Fanuc KAREL source: kt00489.KL

-- PROVISIONAL review KL for V1013-1; original PC SHA256 af2217d419cc08992401e6106b01a0b923f42a5de7de44bf260eaf8e4cc73e97
-- Incomplete behavior may be omitted. Consult companion uncertainty JSON. Do not deploy.
PROGRAM KT00489
%NOLOCKGROUP
-- UNRESOLVED_DECL P1 type=000101
-- UNRESOLVED_DECL P2 type=000199
-- UNRESOLVED_DECL OUT type=000101
BEGIN
  -- UNRESOLVED_PC offsets 5-34; opcodes 49,49,7E,60,4A
  -- UNRESOLVED_PC offsets 39-43; opcodes 7F
END KT00489
